Staubli VAL3: updateJointPos.pgx

program updateJointPos(num x_nIndex)
  local jointRx l_jRef
  local pointRx l_pPos
  local tool l_tTool
  local jointRx l_jResult
begin
  // 回退前，基于后一个点[x_nIndex+1]或当前位置，重新更新jPointRec[x_nIndex]
  if bFirstUpdate==true
    l_jRef=herej()
  else
    // 参考关节l_jRef选择[x_nIndex+1]点
    if nMoveTypeRec[x_nIndex+1]==3
      l_jRef=jPointRec[x_nIndex+1,0]
    else
      l_jRef=jPointRec[x_nIndex+1,1]
    endIf
  endIf
  //
  // update joint
  link(l_tTool,flange)
  l_tTool.trsf=trToolRec[x_nIndex]
  l_pPos=jointToPoint(l_tTool,world,jPointRec[x_nIndex,1])
  pointToJoint(l_tTool,l_jRef,l_pPos,l_jResult)
  if jPointRec[x_nIndex,1]!=l_jResult
    jPointRec[x_nIndex,1]=l_jResult
    logMsg("更新jPointRec["+toString("",x_nIndex)+",1]")
  endIf
  // Movec have two points
  if nMoveTypeRec[x_nIndex]==3
    l_pPos=jointToPoint(l_tTool,world,jPointRec[x_nIndex,0])
    pointToJoint(l_tTool,jPointRec[x_nIndex,1],l_pPos,l_jResult)
    if jPointRec[x_nIndex,0]!=l_jResult
      jPointRec[x_nIndex,0]=l_jResult
      logMsg("更新jPointRec["+toString("",x_nIndex)+",0]")
    endIf
  endIf
end
